{attribute 'qualified_only'}
{attribute 'strict'}
TYPE E_SystemState :
(
	Start 	:= 0,
	Stop 	:= 1,
	Reset	:= 2,
	Fault	:= 99
) INT;
END_TYPE

(* stored: Version 1.1.0.1
   DUT E_SystemState: Id {814ed138-9d9b-47bc-a7e4-af06d745d16d} *)
